FUNCTION_BLOCK T_SafeOpMode_Tests EXTENDS TcUnit.FB_TestSuite
VAR
    // Test_ExactlyOneInputSelectsOutput
    group_1 : T_SafeGroup;
    fb_1 : T_SafeOpMode(group := group_1);
    // Test_ConnectedRestartRequiresRestartSequence
    group_2 : T_SafeGroup;
    fb_2 : T_SafeOpMode(group := group_2);
    // Test_SlowModeChangeGivesDiscrepancyError
    group_3 : T_SafeGroup;
    fb_3 : T_SafeOpMode(group := group_3) := (Parameters := (DiscrepancyTime := T#100MS));
    state_3 : INT := 10;
    waitTimer_3 : TON;
    // Test_OneConnectedInputIsRefused
    group_4 : T_SafeGroup;
    fb_4 : T_SafeOpMode(group := group_4);
END_VAR

Test_ExactlyOneInputSelectsOutput();
Test_ConnectedRestartRequiresRestartSequence();
Test_SlowModeChangeGivesDiscrepancyError();
Test_OneConnectedInputIsRefused();

METHOD PRIVATE Test_ConnectedRestartRequiresRestartSequence
TcUnit.TEST(__POUNAME());
// act
group_2(Run := TRUE);
fb_2(Restart := FALSE, OpIn1 := TRUE, OpIn2 := FALSE);
group_2(Run := TRUE);
fb_2(Restart := FALSE, OpIn1 := TRUE, OpIn2 := FALSE);
// assert
AssertEquals_BOOL(Expected := FALSE, Actual := fb_2.OpOut1, Message := 'no output before restart');
group_2(Run := TRUE);
fb_2(Restart := TRUE, OpIn1 := TRUE, OpIn2 := FALSE);
AssertEquals_BYTE(Expected := TO_BYTE(E_SafeFbState.Start), Actual := fb_2.State, Message := 'state START while restart held');
group_2(Run := TRUE);
fb_2(Restart := FALSE, OpIn1 := TRUE, OpIn2 := FALSE);
AssertEquals_BOOL(Expected := TRUE, Actual := fb_2.OpOut1, Message := 'output on after restart falling edge');
TEST_FINISHED_NAMED(__POUNAME());
END_METHOD

METHOD PRIVATE Test_ExactlyOneInputSelectsOutput
TcUnit.TEST(__POUNAME());
// act: STOP -> SAFE -> RUN (no Restart connected: automatic)
group_1(Run := TRUE);
fb_1(OpIn1 := FALSE, OpIn2 := TRUE);
group_1(Run := TRUE);
fb_1(OpIn1 := FALSE, OpIn2 := TRUE);
// assert
AssertEquals_BOOL(Expected := TRUE, Actual := fb_1.OpOut2, Message := 'selected mode output on');
AssertEquals_BOOL(Expected := FALSE, Actual := fb_1.OpOut1, Message := 'other outputs off');
AssertEquals_BYTE(Expected := TO_BYTE(E_SafeFbState.Run), Actual := fb_1.State, Message := 'state RUN');
// act: second input also set
group_1(Run := TRUE);
fb_1(OpIn1 := TRUE, OpIn2 := TRUE);
AssertEquals_BOOL(Expected := FALSE, Actual := fb_1.OpOut2, Message := 'all outputs off with two modes selected');
AssertEquals_BYTE(Expected := TO_BYTE(E_SafeFbState.Safe), Actual := fb_1.State, Message := 'state SAFE');
TEST_FINISHED_NAMED(__POUNAME());
END_METHOD

METHOD PRIVATE Test_SlowModeChangeGivesDiscrepancyError
TcUnit.TEST(__POUNAME());
waitTimer_3();

CASE state_3 OF
    10:
        // arrange: mode 1 selected and running
        group_3(Run := TRUE);
        fb_3(OpIn1 := TRUE, OpIn2 := FALSE);
        group_3(Run := TRUE);
        fb_3(OpIn1 := TRUE, OpIn2 := FALSE);
        state_3 := 20;
        waitTimer_3(IN := TRUE, PT := T#250MS);
    20:
        // act: leave mode 1 without selecting another
        group_3(Run := TRUE);
        fb_3(OpIn1 := FALSE, OpIn2 := FALSE);

        IF NOT waitTimer_3.Q THEN
            RETURN;
        END_IF

        waitTimer_3(IN := FALSE);
        // assert
        AssertEquals_BOOL(Expected := TRUE, Actual := fb_3.Error, Message := 'discrepancy error after time without a mode');
        AssertEquals_BYTE(Expected := TO_BYTE(E_SafeFbState.Error), Actual := fb_3.State, Message := 'state ERROR');
        AssertEquals_WORD(Expected := WORD#1, Actual := fb_3.Diag, Message := 'diag bit 0');
        TEST_FINISHED_NAMED(__POUNAME());
        state_3 := 10;
END_CASE
END_METHOD

METHOD PRIVATE Test_OneConnectedInputIsRefused
TcUnit.TEST(__POUNAME());
// arrange / act: OpIn1 is the only connected input, which the Safety Editor refuses
group_4(Run := TRUE);
fb_4(OpIn1 := TRUE);
group_4(Run := TRUE);
fb_4(OpIn1 := TRUE);
// assert
AssertEquals_BOOL(Expected := TRUE, Actual := fb_4.Error, Message := 'configuration error reported');
AssertEquals_BYTE(Expected := TO_BYTE(E_SafeFbState.Error), Actual := fb_4.State, Message := 'state ERROR');
AssertEquals_WORD(Expected := WORD#16#8000, Actual := fb_4.Diag, Message := 'diag bit 15 configuration refused');
AssertEquals_BOOL(Expected := FALSE, Actual := fb_4.OpOut1, Message := 'OpOut1 stays at its safe value');
AssertEquals_BOOL(Expected := TRUE, Actual := group_4.FbErr, Message := 'the group sees an FB error');
// act: ErrAck 0 -> 1 -> 0 does not clear a configuration error
group_4(Run := TRUE, ErrAck := TRUE);
fb_4(OpIn1 := TRUE);
group_4(Run := TRUE, ErrAck := TRUE);
fb_4(OpIn1 := TRUE);
group_4(Run := TRUE, ErrAck := FALSE);
fb_4(OpIn1 := TRUE);
AssertEquals_BOOL(Expected := TRUE, Actual := fb_4.Error, Message := 'error not acknowledged');
AssertEquals_WORD(Expected := WORD#16#8000, Actual := fb_4.Diag, Message := 'diag bit 15 kept');
TEST_FINISHED_NAMED(__POUNAME());
END_METHOD

END_FUNCTION_BLOCK

(* stored: Version 1.1.0.1
   POU T_SafeOpMode_Tests: Id {d0130fc1-9d06-5052-9dad-6e22ca0784de}, SpecialFunc None
   Method Test_ConnectedRestartRequiresRestartSequence: Id {f740a1ec-4a81-5461-a63f-89e5adc985f1}
   Method Test_ExactlyOneInputSelectsOutput: Id {3b990399-42cf-5606-b314-eec448d34948}
   Method Test_SlowModeChangeGivesDiscrepancyError: Id {77cb4e41-82ca-565a-b75f-291378702b4f}
   Method Test_OneConnectedInputIsRefused: Id {8c241beb-1510-4f54-b648-73f089e43615} *)
